Staubli VAL3: Trsf2Matrix.pgx

public program Trsf2Matrix(trsf x_trTrsf, num& x_nMatrix[] (dimensions=2))
  local num ax
  local num ay
  local num az
  local num nx
  local num ny
  local num nz
  local num ox
  local num oy
  local num oz
  local num px
  local num py
  local num pz
  local num rx
  local num ry
  local num rz
  local num x
  local num y
  local num z
begin
  //Trsf转换成Matrik
  x=x_trTrsf.x
  y=x_trTrsf.y
  z=x_trTrsf.z
  rx=x_trTrsf.rx
  ry=x_trTrsf.ry
  rz=x_trTrsf.rz
  //
  nx=cos(ry)*cos(rz)
  ny=sin(rx)*sin(ry)*cos(rz)+cos(rx)*sin(rz)
  nz=-cos(rx)*sin(ry)*cos(rz)+sin(rx)*sin(rz)
  ox=-cos(ry)*sin(rz)
  oy=-sin(rx)*sin(ry)*sin(rz)+cos(rx)*cos(rz)
  oz=cos(rx)*sin(ry)*sin(rz)+sin(rx)*cos(rz)
  ax=sin(ry)
  ay=-sin(rx)*cos(ry)
  az=cos(rx)*cos(ry)
  px=x
  py=y
  pz=z
  //
  x_nMatrix[0,0]=nx
  x_nMatrix[0,1]=ny
  x_nMatrix[0,2]=nz
  x_nMatrix[0,3]=0
  x_nMatrix[1,0]=ox
  x_nMatrix[1,1]=oy
  x_nMatrix[1,2]=oz
  x_nMatrix[1,3]=0
  x_nMatrix[2,0]=ax
  x_nMatrix[2,1]=ay
  x_nMatrix[2,2]=az
  x_nMatrix[2,3]=0
  x_nMatrix[3,0]=px
  x_nMatrix[3,1]=py
  x_nMatrix[3,2]=pz
  x_nMatrix[3,3]=1
end
